(* IEC 61131-3 sources: JingjiangMoonbox/Application/Application/任务列表/TensionTask/张力控制/收放料/翻转架补偿, 6 files *)

(* ---- KS_CalcFilmLenth_TowerToNextRoller.st ---- *)
(*@CES
Name=KS_CalcFilmLenth_TowerToNextRoller
Type=FunctionBlock
TypeGuid=6f9dac99-8de1-4efc-8465-68ac443b7d08
Guid=4de748ae-c124-4dda-9073-dd74e9313ddf
HasDeclaration=True
HasImplementation=True
*)
{DECLARATION}
FUNCTION KS_CalcFilmLenth_TowerToNextRoller : INT(*计算放料架到第一个辊之间的料长*)
VAR_INPUT
(*	i_xDir_Rev:BOOL;(*方向取反|默认翻转架运动和绝对值位置变化方向一致|逆时针转动为正方向。*)*)
	i_dwAbsPos_0Rad:DWORD;(*写入0弧度对应的绝对值位置*)
	i_dwAbsPos_Cur:DWORD;(*当前绝对位置*)

	i_iTime_PlcCycle:INT:=20;
	i_rDiam_CurAxis:REAL;(*当前卷径|直径mm*)
	i_rDiam_Tower:REAL;(*翻转架直径mm*)
	i_rDiam_NextRoller:REAL;(*翻转架后第一个导辊直径mm*)

	i_rXPos_NextRoller:REAL;(*mm*)
	i_rYPos_NextRoller:REAL;(*mm*)
	i_lrTheta_Cur:LREAL;(*当前弧度值*)
	i_lrLastTheta:LREAL;(*上个周期的弧度值*)
	i_plrDeltaW_RPMIN:POINTER TO LREAL;
	(*2022.5.17.101635*)
	i_rDiam_DeflectorRollPos:REAL;(*翻料架的导向辊圆心运动直径|距离翻转架圆心=该值/2|mm*)
	i_rDiam_DeflectorRoller:REAL;(*翻料架上导向辊的直径|mm*)
	i_xFilmTouchRoller:BOOL;(*料膜接触到导向辊标志*)
	i_byMaterialPath:BYTE;(*材料行走路径|0:料膜和下个辊外公切线走料
										 1:料膜和下个辊内公切线走料
							PS:放料上裁刀i_byMaterialPath=0
							   放料下裁刀i_byMaterialPath=1
							   收料上裁刀i_byMaterialPath=0
							   收料下裁刀i_byMaterialPath=1*)
END_VAR
VAR
	lrTemp:LREAL;
	lrTemp1:LREAL;
	lrC: LREAL;
	lrts: LREAL;(*采样周期|s*)
	lrRadius_CurAxis:LREAL;(*当前轴半径|m*)
	lrRadius_Tower: LREAL;(*翻转架半径|M*)
	lrRadius_NextRoller: LREAL;(*下个导辊的半径|M*)
	lrX_NextRoller: LREAL;(*下个辊的x位置|m*)
	lrY_NextRoller: LREAL;(*下个辊的Y位置|m*)
	lrRadius_DeflectorRollPos:LREAL;(*翻料架的导向辊圆心运动半径|距离翻转架圆心=该值/2|m*)
	lrRadius_DeflectorRoller:LREAL;(*翻料架上导向辊的半径|m*)
	dwAbsPos_0Rad: DWORD;(*写入0弧度对应的绝对值位置*)
	lrTheta_Cur: LREAL;(*当前弧度*)
	lrPi:LREAL:=3.1415926;
(*	dwAbsPos_Cycle:DWORD:=131072;*)
	iErr: INT;
	lrDeltFilmLen: LREAL;
	lrLastTheta_Cur: LREAL;
	lrDeltW: LREAL;
	lrDeltW_RPMIN: LREAL;
END_VAR
{IMPLEMENTATION}
dwAbsPos_0Rad:=i_dwAbsPos_0Rad;
lrLastTheta_Cur:=i_lrLastTheta;
lrTheta_Cur:=i_lrTheta_Cur;

(*根据手册公式实现*)
(*根据手册单位进行对应转换*)
lrts:=INT_TO_LREAL(i_iTime_PlcCycle)/1000;
lrRadius_CurAxis:=i_rDiam_CurAxis/1000/2;
lrRadius_Tower:=i_rDiam_Tower/1000/2;
lrRadius_NextRoller:=i_rDiam_NextRoller/1000/2;
lrX_NextRoller:=i_rXPos_NextRoller/1000;
lrY_NextRoller:=i_rYPos_NextRoller/1000;
lrRadius_DeflectorRollPos:=i_rDiam_DeflectorRollPos/1000/2;
lrRadius_DeflectorRoller:=i_rDiam_DeflectorRoller/1000/2;

(*lrC的计算不考虑内切还是外切都是按照外切计算长度|两种的变化率保持一致*)
IF NOT i_xFilmTouchRoller THEN(*未接触到导向辊|*)
	lrC:=lrX_NextRoller*lrX_NextRoller+lrY_NextRoller*lrY_NextRoller+
		lrRadius_Tower*lrRadius_Tower-
		lrRadius_NextRoller*lrRadius_NextRoller-
		lrRadius_CurAxis*lrRadius_CurAxis+
		2*lrRadius_NextRoller*lrRadius_CurAxis;
ELSE(*接触到导向辊*)
	lrC:=lrX_NextRoller*lrX_NextRoller+lrY_NextRoller*lrY_NextRoller+
		lrRadius_DeflectorRollPos*lrRadius_DeflectorRollPos+
		2*lrRadius_DeflectorRoller*lrRadius_NextRoller-
		lrRadius_DeflectorRoller*lrRadius_DeflectorRoller-
		lrRadius_NextRoller*lrRadius_NextRoller;
END_IF
IF lrC<=0 THEN
	iErr:=-1;
END_IF

IF iErr=0 THEN
	CASE i_byMaterialPath OF
		1:(*内公切线走料|下裁刀方式*)
			IF NOT i_xFilmTouchRoller THEN(*未接触到导向辊|公式和外公切线使用同样的公式*)
				lrTemp:=lrC-2*lrRadius_Tower*(lrX_NextRoller*COS(lrTheta_Cur)+lrY_NextRoller*SIN(lrTheta_Cur));
				lrTemp1:=lrC-2*lrRadius_Tower*(lrX_NextRoller*COS(lrLastTheta_Cur)+lrY_NextRoller*SIN(lrLastTheta_Cur));
			ELSE(*接触到导向辊*)
				lrTemp:=lrC+2*lrRadius_DeflectorRollPos*(lrX_NextRoller*SIN(lrTheta_Cur)-lrY_NextRoller*COS(lrTheta_Cur));
				lrTemp1:=lrC+2*lrRadius_DeflectorRollPos*(lrX_NextRoller*SIN(lrLastTheta_Cur)-lrY_NextRoller*COS(lrLastTheta_Cur));
			END_IF
	ELSE(*外公切线走料|上裁刀方式*)
		IF NOT i_xFilmTouchRoller THEN(*未接触到导向辊|*)
			lrTemp:=lrC-2*lrRadius_Tower*(lrX_NextRoller*COS(lrTheta_Cur)+lrY_NextRoller*SIN(lrTheta_Cur));
			lrTemp1:=lrC-2*lrRadius_Tower*(lrX_NextRoller*COS(lrLastTheta_Cur)+lrY_NextRoller*SIN(lrLastTheta_Cur));
		ELSE(*接触到导向辊*)
			lrTemp:=lrC-2*lrRadius_DeflectorRollPos*(lrX_NextRoller*SIN(lrTheta_Cur)-lrY_NextRoller*COS(lrTheta_Cur));
			lrTemp1:=lrC-2*lrRadius_DeflectorRollPos*(lrX_NextRoller*SIN(lrLastTheta_Cur)-lrY_NextRoller*COS(lrLastTheta_Cur));
		END_IF
	END_CASE

	IF lrTemp>=0 THEN
		lrTemp:=SQRT(lrTemp);
	ELSE
		iErr:=-2;
	END_IF

	IF lrTemp1>=0 THEN
		lrTemp1:=SQRT(lrTemp1);
	ELSE
		iErr:=-3;
	END_IF

	IF iErr=0 THEN
		lrDeltFilmLen:=lrTemp-lrTemp1;
	END_IF

	IF lrRadius_CurAxis<>0 THEN
		lrDeltW:=lrDeltFilmLen/lrts/lrRadius_CurAxis;
	END_IF

	lrDeltW_RPMIN:=lrDeltW*60/2/lrPi;
END_IF

IF i_plrDeltaW_RPMIN<>0 THEN
	i_plrDeltaW_RPMIN^:=lrDeltW_RPMIN;
END_IF

KS_CalcFilmLenth_TowerToNextRoller:=iErr;

(* ---- KS_CalcRadByAbsEnc.st ---- *)
(*@CES
Name=KS_CalcRadByAbsEnc
Type=FunctionBlock
TypeGuid=6f9dac99-8de1-4efc-8465-68ac443b7d08
Guid=0e1ec2d5-a158-4810-bac7-8538ad8533d7
HasDeclaration=True
HasImplementation=True
*)
{DECLARATION}
FUNCTION KS_CalcRadByAbsEnc : LREAL(*返回当前弧度|需要标定0弧度对应的绝对位置值*)
VAR_INPUT
	i_xDir_Rev:BOOL;(*方向取反|默认翻转架运动和绝对值位置变化方向一致|逆时针转动为正方向。*)
	i_dwAbsPos_0Rad:DWORD;(*0弧度对应的绝对值位置*)
	i_dwAbsPos_Cur:DWORD;(*当前绝对位置*)
	i_dwAbsPos_Cycle:DWORD:=131072;(*编码器线束*)
END_VAR
VAR
	dwTemp:DWORD;
	lrTemp:LREAL;
	dwAbsPos_Cycle:DWORD;
	lrTheta_Cur: LREAL;
END_VAR
{IMPLEMENTATION}
dwAbsPos_Cycle:=i_dwAbsPos_Cycle;
dwTemp:=(i_dwAbsPos_Cur+dwAbsPos_Cycle-i_dwAbsPos_0Rad) MOD (dwAbsPos_Cycle);
IF dwAbsPos_Cycle<>0 THEN
	lrTemp:=2*gc_lrPI/dwAbsPos_Cycle*dwTemp;(*变化的角度*)
END_IF

IF i_xDir_Rev THEN
	lrTemp:=-lrTemp;
END_IF

lrTheta_Cur:=lrTemp;
IF lrTemp>2*gc_lrPI THEN
	lrTheta_Cur:=lrTemp-2*gc_lrPI;
ELSIF lrTemp<0 THEN
	lrTheta_Cur:=lrTemp+2*gc_lrPI;
END_IF

KS_CalcRadByAbsEnc:=lrTheta_Cur;

(* ---- KS_FilmToTowerRollerDis.st ---- *)
(*@CES
Name=KS_FilmToTowerRollerDis
Type=FunctionBlock
TypeGuid=6f9dac99-8de1-4efc-8465-68ac443b7d08
Guid=026cf6eb-c0d8-494e-aced-39e104fa3684
HasDeclaration=True
HasImplementation=True
*)
{DECLARATION}
FUNCTION KS_FilmToTowerRollerDis : INT(*计算料膜到翻料架导向辊的距离|负值代表错误*)
VAR_INPUT
	i_byMaterialPath:BYTE;(*材料行走路径|0:料膜和下个辊外公切线走料
										 1:料膜和下个辊内公切线走料
							PS:放料上裁刀i_byMaterialPath=0
							   放料下裁刀i_byMaterialPath=1
							   收料上裁刀i_byMaterialPath=0
							   收料下裁刀i_byMaterialPath=1*)
	i_rDiam_DeflectorRollPos:REAL;(*翻料架的导向辊圆心运动直径|距离翻转架圆心=该值/2|mm*)
	i_rDiam_DeflectorRoller:REAL;(*翻料架上导向辊的直径|mm*)
	i_rDiam_CurAxis:REAL;(*当前卷径|直径mm*)
	i_rDiam_Tower:REAL;(*翻转架直径mm*)
	i_rDiam_NextRoller:REAL;(*翻转架后第一个导辊直径mm*)
	i_rXPos_NextRoller:REAL;(*mm*)
	i_rYPos_NextRoller:REAL;(*mm*)
	i_lrTheta_Cur:LREAL;(*当前弧度值*)
	i_prFilmToTowerRollerDis:POINTER TO REAL;(*mm*)
	i_pxFilmTouchRoller:POINTER TO BOOL;(**)
END_VAR
VAR
	iRtn: INT;
	lrRadius_DeflectorRollPos:LREAL;(*翻料架的导向辊圆心运动半径|距离翻转架圆心=该值/2|m*)
	lrRadius_DeflectorRoller:LREAL;(*翻料架上导向辊的直径|m*)
	lrRadius_CurAxis:LREAL;(*当前轴半径|m*)
	lrRadius_Tower: LREAL;(*翻转架半径|M*)
	lrRadius_NextRoller: LREAL;(*下个导辊的半径|M*)
	lrX_NextRoller: LREAL;(*下个辊的x位置|m*)
	lrY_NextRoller: LREAL;(*下个辊的Y位置|m*)
	lrTheta_Cur: LREAL;(*当前弧度*)
	lrFilmToTowerRollerDis:LREAL;
	lrIy: LREAL;
	lrIx: LREAL;
	lrUx: LREAL;
	lrUy: LREAL;
	lrDelta: LREAL;
	lrp1: LREAL;
	lrp2: LREAL;
	lrq: LREAL;
	lrA: LREAL;
	lrB: LREAL;
	lrC: LREAL;
	lrD: LREAL;
	lrD0: LREAL;
	lrD1: LREAL;
	xFilmTouchRoller: BOOL;(*料膜接触到了辊子*)
END_VAR
{IMPLEMENTATION}
(*计算公式:
Ix、Iy-导向辊的坐标 Ix=i_rDiam_DeflectorRollPos/2*SIN(i_rTheta_Cur)；
				    Iy=-i_rDiam_DeflectorRollPos/2*Cos(i_rTheta_Cur);
Ux、Uy当前轴的坐标 Ux=i_rDiam_Tower/2*Cos(i_rTheta_Cur);
				   Uy=i_rDiam_Tower/2*Sin(i_rTheta_Cur);
计算启动启动的条件为Ux<Ix;
Delta=(Ux-i_rXPos_NextRoller)^2+(Uy-i_rYPos_NextRoller)^2-(i_rDiam_CurAxis-i_rDiam_NextRoller)^2/4;
P1=i_rDiam_CurAxis/2*(i_rXPos_NextRoller^2+i_rYPos_NextRoller^2-i_rXPos_NextRoller*Ux-i_rYPos_NextRoller*Uy);
P2=i_rDiam_NextRoller/2*(Ux^2+Uy^2-i_rXPos_NextRoller*Ux-i_rYPos_NextRoller*Uy);
q=Ux*i_rYPos_NextRoller-Uy*i_rXPos_NextRoller;
A=(i_rXPos_NextRoller-Ux)*(i_rDiam_CurAxis-i_rDiam_NextRoller)/2+(Uy-i_rYPos_NextRoller)*SQRT(Delta);
B=(i_rYPos_NextRoller-Uy)*(i_rDiam_CurAxis-i_rDiam_NextRoller)/2+(i_rXPos_NextRoller-Ux)*SQRT(Delta);
C=-P1-P2+q*SQRT(Delta);
D0=A*Ix+B*Iy+C;
D=D0/SQRT(A^2+B^2);
*)
IF i_pxFilmTouchRoller<>0 THEN
	xFilmTouchRoller:=i_pxFilmTouchRoller^;
END_IF

lrRadius_CurAxis:=i_rDiam_CurAxis/1000/2;
lrRadius_Tower:=i_rDiam_Tower/1000/2;
lrRadius_NextRoller:=i_rDiam_NextRoller/1000/2;
lrX_NextRoller:=i_rXPos_NextRoller/1000;
lrY_NextRoller:=i_rYPos_NextRoller/1000;
lrRadius_DeflectorRollPos:=i_rDiam_DeflectorRollPos/1000/2;
lrRadius_DeflectorRoller:=i_rDiam_DeflectorRoller/1000/2;
lrTheta_Cur:=i_lrTheta_Cur;
lrFilmToTowerRollerDis:=0;

CASE i_byMaterialPath OF
	1:(*内公切线|D是正值代表远离-下裁刀方式*)
		(*计算导向辊的坐标*)
		lrIx:=-lrRadius_DeflectorRollPos*SIN(lrTheta_Cur);
		lrIy:=lrRadius_DeflectorRollPos*COS(lrTheta_Cur);
		(*计算当前轴的坐标*)
		lrUx:=lrRadius_Tower*COS(lrTheta_Cur);
		lrUy:=lrRadius_Tower*SIN(lrTheta_Cur);
		IF lrUx < lrIx THEN(*启动计算*)
			lrDelta:=EXPT((lrUx-lrX_NextRoller),2)+EXPT((lrUy-lrY_NextRoller),2)-EXPT((lrRadius_CurAxis+lrRadius_NextRoller),2);
			IF lrDelta>=0 THEN
				lrp1:=lrRadius_CurAxis*(EXPT(lrX_NextRoller,2)+EXPT(lrY_NextRoller,2)-lrX_NextRoller*lrUx-lrY_NextRoller*lrUy);
				lrp2:=lrRadius_NextRoller*(EXPT(lrUx,2)+EXPT(lrUy,2)-lrX_NextRoller*lrUx-lrY_NextRoller*lrUy);
				lrq:=lrUx*lrY_NextRoller-lrUy*lrX_NextRoller;
				lrA:=(lrX_NextRoller-lrUx)*(lrRadius_CurAxis+lrRadius_NextRoller)-(lrUy-lrY_NextRoller)*SQRT(lrDelta);
				lrB:=(lrY_NextRoller-lrUy)*(lrRadius_CurAxis+lrRadius_NextRoller)-(lrX_NextRoller-lrUx)*SQRT(lrDelta);
				lrC:=-lrp1+lrp2-lrq*SQRT(lrDelta);
				lrD0:=lrA*lrIx+lrB*lrIy+lrC;
				lrD1:=EXPT(lrA,2)+EXPT(lrB,2);
				IF lrD1>0 THEN
					lrD:=(lrD0)/SQRT(lrD1);(*m*)
				ELSE
					iRtn:=-3;
				END_IF
			ELSE
				iRtn:=-2;
			END_IF
		ELSE
			iRtn:=-1;
		END_IF
ELSE(*外公切线|D是负值代表远离-上裁刀方式*)
		(*计算导向辊的坐标*)
		lrIx:=lrRadius_DeflectorRollPos*SIN(lrTheta_Cur);
		lrIy:=-lrRadius_DeflectorRollPos*COS(lrTheta_Cur);
		(*计算当前轴的坐标*)
		lrUx:=lrRadius_Tower*COS(lrTheta_Cur);
		lrUy:=lrRadius_Tower*SIN(lrTheta_Cur);
		IF lrUx < lrIx THEN(*启动计算*)
			lrDelta:=EXPT((lrUx-lrX_NextRoller),2)+EXPT((lrUy-lrY_NextRoller),2)-EXPT((lrRadius_CurAxis-lrRadius_NextRoller),2);
			IF lrDelta>=0 THEN
				lrp1:=lrRadius_CurAxis*(EXPT(lrX_NextRoller,2)+EXPT(lrY_NextRoller,2)-lrX_NextRoller*lrUx-lrY_NextRoller*lrUy);
				lrp2:=lrRadius_NextRoller*(EXPT(lrUx,2)+EXPT(lrUy,2)-lrX_NextRoller*lrUx-lrY_NextRoller*lrUy);
				lrq:=lrUx*lrY_NextRoller-lrUy*lrX_NextRoller;
				lrA:=(lrX_NextRoller-lrUx)*(lrRadius_CurAxis-lrRadius_NextRoller)+(lrUy-lrY_NextRoller)*SQRT(lrDelta);
				lrB:=(lrY_NextRoller-lrUy)*(lrRadius_CurAxis-lrRadius_NextRoller)+(lrX_NextRoller-lrUx)*SQRT(lrDelta);
				lrC:=-lrp1-lrp2+lrq*SQRT(lrDelta);
				lrD0:=lrA*lrIx+lrB*lrIy+lrC;
				lrD1:=EXPT(lrA,2)+EXPT(lrB,2);
				IF lrD1>0 THEN
					lrD:=(lrD0)/SQRT(lrD1);(*m*)
				ELSE
					iRtn:=-3;
				END_IF
			ELSE
				iRtn:=-2;
			END_IF
		ELSE
			iRtn:=-1;
		END_IF
END_CASE

IF iRtn=0 THEN(*算出来了*)
	(*增加了0.01M的回差*)
	IF NOT xFilmTouchRoller THEN
		IF lrD+lrRadius_DeflectorRoller>=0 THEN
			xFilmTouchRoller:=TRUE;
		END_IF
	ELSIF lrD+lrRadius_DeflectorRoller<-0.01 THEN
		xFilmTouchRoller:=FALSE;
	END_IF
ELSE
	xFilmTouchRoller:=FALSE;
END_IF

IF i_pxFilmTouchRoller<>0 THEN
	i_pxFilmTouchRoller^:=xFilmTouchRoller;
END_IF

IF i_prFilmToTowerRollerDis<>0 THEN
	i_prFilmToTowerRollerDis^:=LREAL_TO_REAL(lrD*1000.0);
END_IF
KS_FilmToTowerRollerDis:=iRtn;

(* ---- KS_GetAbsPos_0Rad.st ---- *)
(*@CES
Name=KS_GetAbsPos_0Rad
Type=FunctionBlock
TypeGuid=6f9dac99-8de1-4efc-8465-68ac443b7d08
Guid=6804038e-cb39-41e6-bf94-3a2690a56994
HasDeclaration=True
HasImplementation=True
*)
{DECLARATION}
FUNCTION KS_GetAbsPos_0Rad : DWORD(*获取0弧度对应的*)
VAR_INPUT
	i_xGetAbsPos:BOOL;
	i_dwAbsPos_Cur:DWORD;(*当前绝对位置*)
	i_pdwAbsPos_0Rad:POINTER TO DWORD;(*写入0弧度对应的绝对值位置*)
END_VAR
VAR
END_VAR
{IMPLEMENTATION}
IF i_xGetAbsPos THEN
	IF i_pdwAbsPos_0Rad<>0 THEN
		i_pdwAbsPos_0Rad^:=i_dwAbsPos_Cur;
	END_IF
END_IF

(* ---- KS_FB_FiltByAver.st ---- *)
(*@CES
Name=KS_FB_FiltByAver
Type=FunctionBlock
TypeGuid=6f9dac99-8de1-4efc-8465-68ac443b7d08
Guid=d55a5298-8c05-4803-b072-b92952ba6371
HasDeclaration=True
HasImplementation=True
*)
{DECLARATION}
FUNCTION_BLOCK KS_FB_FiltByAver(*通过平均进行滤波|2020.10.8.140809更新。*)
(*2023.09.04.122927 为了减少空间利用-将最大滤波次数输出由60个修改到了30个|
滤波数组类型LREAL修改为了real*)
VAR_INPUT
	i_xEn					:BOOL;
	i_iFiltTimes			:INT;(*滤波次数，最大60*)
	i_dwDataAdr				:DWORD;(*需要滤波的数据地址*)
	i_byDataType			:TypEnumDataType;(*滤波的数据类型*)
	i_xFrom0Average			:BOOL;(*从0开始滤波@2024.05.21.163305*)
END_VAR
VAR_OUTPUT
	o_xEn					:BOOL;
(*	o_alrArrData			:ARRAY [1..60] OF LREAL;(*存放数据的数组，1是最新数据*)*)
	o_alrArrData			:ARRAY [1..30] OF LREAL;(*存放数据的数组，1是最新数据@2023.09.04.123126*)
	o_rFiltData			:REAL;(*滤波后的值*)
	o_iCode					:INT;
END_VAR
VAR
	plrData				:POINTER TO LREAL;
	prData				:POINTER TO REAL;
	pdiData				:POINTER TO DINT;
	pdwData				:POINTER TO DWORD;
	piData				:POINTER TO INT;
	pwData				:POINTER TO WORD;
	pbyData				:POINTER TO BYTE;
	pxData				:POINTER TO BOOL;

	lrData				:LREAL;(*进行滤波的数据*)
	iN					:INT;
	lrDataSum			:LREAL;(**)
	xArrInit			:BOOL;(*滤波数组初始化*)
	iInitCnt			:INT:=0;
	iPreFiltTimes		:INT;
	xPreFilterTimeInit	:BOOL:=FALSE;
END_VAR
{IMPLEMENTATION}
IF i_iFiltTimes>30 THEN i_iFiltTimes:=30;ELSIF i_iFiltTimes<=0 THEN i_iFiltTimes:=1;END_IF
o_xEn:=i_xEn;
IF NOT xPreFilterTimeInit THEN
	xPreFilterTimeInit:=TRUE;
	iPreFiltTimes:=i_iFiltTimes;
END_IF

plrData:=0;
plrData:=0;
prData:=0;
pdiData:=0;
pdwData:=0;
piData:=0;
pwData:=0;
pbyData:=0;
pxData:=0;
lrData:=0;
o_iCode:=0;
IF i_dwDataAdr<>0 THEN(*数据地址有效了 我们可以进行滤波*)
	CASE i_byDataType OF
	TYPE_LREAL:
		plrData:=i_dwDataAdr;
		lrData:=plrData^;
	TYPE_REAL:
		prData:=i_dwDataAdr;
		lrData:=REAL_TO_LREAL(prData^);
	TYPE_DINT:
		pdiData:=i_dwDataAdr;
		lrData:=DINT_TO_LREAL(pdiData^);
	TYPE_DWORD:
		pdwData:=i_dwDataAdr;
		lrData:=DWORD_TO_LREAL(pdwData^);
	TYPE_INT:
		piData:=i_dwDataAdr;
		lrData:=INT_TO_LREAL(piData^);
	TYPE_WORD:
		pwData:=i_dwDataAdr;
		lrData:=WORD_TO_LREAL(pwData^);
	TYPE_BYTE:
		pbyData:=i_dwDataAdr;
		lrData:=BYTE_TO_LREAL(pbyData^);
	TYPE_BOOL:
		pxData:=i_dwDataAdr;
		lrData:=BOOL_TO_LREAL(pxData^);
	ELSE
		o_iCode:=-2;
	END_CASE
ELSE
	o_iCode:=-1;
	RETURN;
END_IF

IF i_xEn THEN(*滤波使能*)
	IF i_iFiltTimes>iPreFiltTimes THEN(*滤波次数加大了 我们重新初始化数组*)
		xArrInit:=FALSE;
	ELSIF i_iFiltTimes<iPreFiltTimes THEN(*次数减小了 我们只更新数组初始计数值*)
		IF	xArrInit THEN
			iInitCnt:=i_iFiltTimes;
		END_IF
	END_IF

	IF NOT xArrInit THEN(*滤波数组初始化*)
	(*	iInitCnt:=iInitCnt+1;
		IF iInitCnt>=i_iFiltTimes THEN
			xArrInit:=TRUE;
		END_IF
*)		(*滤波初始化时，数据数组一次写入*)
		FOR iN:=1 TO i_iFiltTimes BY 1 DO
			IF i_xFrom0Average THEN
				o_alrArrData[iN]:=0;
			ELSE
				o_alrArrData[iN]:=lrData;
			END_IF
		END_FOR
		xArrInit:=TRUE;
	END_IF

	(*开始进行滤波*)
	IF i_iFiltTimes>=2 THEN
		FOR iN:=i_iFiltTimes TO 2 BY -1 DO
			o_alrArrData[iN]:=o_alrArrData[iN-1];
		END_FOR
	ELSE(*不进行滤波*);
	END_IF
	o_alrArrData[1]:=lrData;

	o_rFiltData:=0;
	IF xArrInit THEN
		lrDataSum:=0;
		FOR	 iN:=1 TO i_iFiltTimes BY 1 DO
			lrDataSum:=lrDataSum+o_alrArrData[iN];
		END_FOR

		o_rFiltData:=LREAL_TO_REAL(lrDataSum/i_iFiltTimes);
	END_IF
ELSE(*不滤波*)
	xArrInit:=FALSE;
	iInitCnt:=0;
	o_rFiltData:=LREAL_TO_REAL(lrData);
END_IF

iPreFiltTimes:=i_iFiltTimes;

(* ---- KS_FB_TowerRadCompensate.st ---- *)
(*@CES
Name=KS_FB_TowerRadCompensate
Type=FunctionBlock
TypeGuid=6f9dac99-8de1-4efc-8465-68ac443b7d08
Guid=99248248-9d66-40a1-9b64-687b8d387c7e
HasDeclaration=True
HasImplementation=True
*)
{DECLARATION}
FUNCTION_BLOCK KS_FB_TowerRadCompensate(*2021.7.26.090725 修改名 增加接口*)
(*2023.6.13.164301 对转速输出增加了10次滤波处理@防止开始时候输出速度抖动*)
(*2023.07.18.094631 翻转架补偿处理最大变化量逻辑中未对过圈问题处理
将滤波次数减小到5次*)
VAR_INPUT
	i_xEn:BOOL;
	i_xAxis_Cur:BOOL;(*当前轴|有效为A轴*)
	i_xConfirmRad:BOOL;
	i_rDiam_CurAxis:REAL;
	i_dwAbsPos_Cur:DWORD;(*当前绝对值位置*)
	i_dwAbsEnCodeResolution:DWORD;(*位置分辨率|131072*)
	(*需要的参数|2021.7.26.090721*)
	I_xTowerDir_Uw:BOOL;(*翻转架和绝对值编码器的方向对应*)
	i_rDiam_Tower:REAL;(*翻转架直径mm*)
	i_rDiam_NextRoller:REAL;(*翻转架后第一个导辊直径mm*)
	i_rXPos_NextRoller:REAL;(*mm*)
	i_rYPos_NextRoller:REAL;(*mm*)
	i_pdwAbsPos_0Rad_AxisA:POINTER TO DWORD;(*A轴0度位置*)
	i_pdwAbsPos_0Rad_AxisB:POINTER TO DWORD;(*B轴0度位置*)
	i_xOnTop:BOOL;(*上下裁刀标志*)
	i_rDiam_DeflectorRollPos:REAL;(*翻料架的导向辊圆心运动直径|距离翻转架圆心=该值/2|mm*)
	i_rDiam_DeflectorRoller:REAL;(*翻料架上导向辊的直径|mm*)
	i_iCycleTime_Plc: INT;
END_VAR
VAR_OUTPUT
	o_rDeltaW_RPMIN: REAL;(*为了不修改外部接口这个变量冲洗定义为了滤波后的值@2023.6.13.163911*)
	o_rTheta_Cur:REAL;(*当前角度*)
	o_rFilmToTowerRollerDis:REAL;(*料膜距离导向辊距离|mm*)
	o_xFilmTouchRoller:BOOL;(*料膜接触到了辊子标志*)
	o_rActDeltaW_RPMIN: REAL;(*当前计算出来的值@2023.6.13.163905*)
END_VAR
VAR
	dwAbsPos_0Rad:DWORD;
	dwAbsPos_Cur:DWORD;
	lrLastTheta:LREAL;
	xInitLastRad:BOOL:=TRUE;
	lrDeltaW_RPMIN:LREAL;(*单个周期的补偿转速*)
	rDiam_CurAxis:REAL;(*放料当前卷径*)
	fbConfirmAbsPos_0Rad: R_TRIG;
	lrTheta_Cur: LREAL;
	lrDeltaTheta_Max: LREAL;
	xCutOnDown: BOOL;(*有效了代表下裁刀*)
	fbKS_FB_FiltByAver: KS_FB_FiltByAver;(*2023.6.13.161714 对当前弧度值进行滤波处理@10次*)
	rDeltaTheta: REAL;		(*2023.07.18.094748*)
END_VAR
{IMPLEMENTATION}
dwAbsPos_Cur:=i_dwAbsPos_Cur;

IF i_xAxis_Cur THEN(*A轴*)
	IF i_pdwAbsPos_0Rad_AxisA<>0 THEN
		dwAbsPos_0Rad:=i_pdwAbsPos_0Rad_AxisA^;
	END_IF
ELSE(*当前轴为B轴*)
	IF i_pdwAbsPos_0Rad_AxisB<>0 THEN
		dwAbsPos_0Rad:=i_pdwAbsPos_0Rad_AxisB^;
	END_IF
END_IF

(*确认0弧度对应的绝对值位置*)
fbConfirmAbsPos_0Rad(CLK:=i_xConfirmRad);
KS_GetAbsPos_0Rad(fbConfirmAbsPos_0Rad.Q, dwAbsPos_Cur, ADR(dwAbsPos_0Rad));
(*当前弧度计算*)
lrTheta_Cur:=KS_CalcRadByAbsEnc(I_xTowerDir_Uw, dwAbsPos_0Rad, dwAbsPos_Cur,i_dwAbsEnCodeResolution );

(*将下面使用的弧度值全部替换为了滤波后的弧度值@2023.6.13.162642*)
(*上个周期弧度值初始化*)
IF i_xConfirmRad OR xInitLastRad THEN(*确认弧度和绝对位置的关系时，重新初始化弧度备份值*)
	fbKS_FB_FiltByAver(i_xEn:= FALSE);(*复位滤波函数*)
	lrLastTheta:=lrTheta_Cur;
END_IF
o_rTheta_Cur:=LREAL_TO_REAL(lrTheta_Cur);
xInitLastRad:=FALSE;

xCutOnDown:=NOT i_xOnTop;

IF i_xEn THEN
	(*2022.5.17.114502 判断是否接触到到导向辊*)
	KS_FilmToTowerRollerDis(
		BOOL_TO_BYTE(xCutOnDown)(*i_byMaterialPath*),
		i_rDiam_DeflectorRollPos(*i_rDiam_DeflectorRollPos*),
		i_rDiam_DeflectorRoller(*i_rDiam_DeflectorRoller*),
		rDiam_CurAxis(*i_rDiam_CurAxis*),
		i_rDiam_Tower(*i_rDiam_Tower*),
		i_rDiam_NextRoller(*i_rDiam_NextRoller*),
		i_rXPos_NextRoller(*i_rXPos_NextRoller*),
		i_rYPos_NextRoller(*i_rYPos_NextRoller*),
		lrTheta_Cur(*i_rTheta_Cur*),
		ADR(o_rFilmToTowerRollerDis)(*i_prFilmToTowerRollerDis*),
		ADR(o_xFilmTouchRoller)(*i_pxFilmTouchRoller*));

	KS_CalcFilmLenth_TowerToNextRoller(
(*		I_xTowerDir_Uw,*)
		dwAbsPos_0Rad,
		dwAbsPos_Cur,
		i_iCycleTime_Plc,
		rDiam_CurAxis,
		i_rDiam_Tower,
		i_rDiam_NextRoller,
		i_rXPos_NextRoller,
		i_rYPos_NextRoller,
		lrTheta_Cur,
		lrLastTheta,
		ADR(lrDeltaW_RPMIN),
		i_rDiam_DeflectorRollPos(*i_rDiam_DeflectorRollPos*),
		i_rDiam_DeflectorRoller(*i_rDiam_DeflectorRoller*),
		o_xFilmTouchRoller(*i_xFilmTouchRoller*),
		BOOL_TO_BYTE(xCutOnDown)(*i_byMaterialPath*));

	(*使能的时候翻转架是在转动的|由于电位器方式时，会有一定时间的死区，该部分
	的处理方式是保持之前的输出转速不变|2021.7.12.174454*)
	(*检查弧度在运动过程中最大的变化量|*)

	(*2023.07.18.094717@过圈问题处理*)
	rDeltaTheta:= LREAL_TO_REAL(ABS(lrTheta_Cur-lrLastTheta));
	IF rDeltaTheta>lrDeltaTheta_Max AND
		rDeltaTheta<gc_lrPI THEN(*2023.07.18.094910  判断过圈*)
		lrDeltaTheta_Max:=rDeltaTheta;
	END_IF
	IF ABS(lrLastTheta-lrTheta_Cur)<lrDeltaTheta_Max/100 THEN(*变化量小于最大的1/100-我们认为进入了电位器电压死区。*)
		(*保持之前的输出量*)
		;(*不更新输出值*)
	ELSE(*正常运动|输出计算值*)
		(*2023.6.13.164033 屏蔽*)
(*		o_lrDeltaW_RPMIN:=lrDeltaW_RPMIN;*)
		o_rActDeltaW_RPMIN:=LREAL_TO_REAL(lrDeltaW_RPMIN);(*修改了变量定义@2023.6.13.164026*)
	END_IF

	(*2023.6.13.163439 对输出的转速进行滤波@不能对输入的角度滤波，过圈会麻烦了*)
	fbKS_FB_FiltByAver(
		i_xEn:= TRUE,
		i_iFiltTimes:=5(*10*),(*滤波时间减小到5个周期*)
		i_dwDataAdr:= ADR(o_rActDeltaW_RPMIN),
		i_byDataType:= TYPE_LREAL,
		i_xFrom0Average:=FALSE,(*2024.05.21.163449*)
		o_xEn=> ,
		o_alrArrData=> ,
		o_rFiltData=> o_rDeltaW_RPMIN,
		o_iCode=> );

	lrLastTheta:=lrTheta_Cur;
ELSE
	xInitLastRad:=TRUE;
	rDiam_CurAxis:=i_rDiam_CurAxis;(*取当前卷径值|在补偿过程中不变化*)
	lrDeltaTheta_Max:=0;
	o_rDeltaW_RPMIN:=0;
	o_rActDeltaW_RPMIN:=0;(*2023.6.13.164229*)
	o_xFilmTouchRoller:=FALSE;
	o_rFilmToTowerRollerDis:=0;
	(*2023.6.13.163637@复位滤波函数*)
	fbKS_FB_FiltByAver(i_xEn:= FALSE);
END_IF

IF i_pdwAbsPos_0Rad_AxisA<>0 AND i_pdwAbsPos_0Rad_AxisB<>0 THEN
	IF i_xAxis_Cur THEN(*A轴*)
		i_pdwAbsPos_0Rad_AxisA^:=dwAbsPos_0Rad;
		IF fbConfirmAbsPos_0Rad.Q THEN(*确认0度值|更新2个轴*)
			(*2个对称*)
			i_pdwAbsPos_0Rad_AxisB^:=(i_dwAbsEnCodeResolution/2+dwAbsPos_0Rad) MOD i_dwAbsEnCodeResolution;
		END_IF
	ELSE(*当前轴为B轴*)
		i_pdwAbsPos_0Rad_AxisB^:=dwAbsPos_0Rad;
		IF fbConfirmAbsPos_0Rad.Q THEN(*确认0度值|更新2个轴*)
			i_pdwAbsPos_0Rad_AxisA^:=(i_dwAbsEnCodeResolution/2+dwAbsPos_0Rad) MOD i_dwAbsEnCodeResolution;
		END_IF
	END_IF
END_IF
